SUBAPPLICATION Softkey_Aux_IXA_TO_Remote_WRITE_BG_Option_OPC (* VT-SoftKey lesen ODER AUX-Zuweisung (Joystick) lesen ODER lokaler Web-Override (z.B. vt-ui-mirror auf demselben Modul) + Remote-OPC-UA-Write an Zielmodul + VT-Hintergrundfarbe (SoftKey UND AUX) aus Remote-Subscribe - Option-Lib- Variante von Softkey_Aux_IXA_TO_Remote_WRITE_BG_OPC: Kommando-Seite komplett inaktiv (echtes INIT_REQ/INIT_CNF, kein VT-Object-Binding) wenn die Option nicht ausgewaehlt ist. Status-Seite (Remote-Subscribe) bleibt unveraendert immer aktiv - reiner Read ohne Seiteneffekt. *)
  (* Standard: 61499-2; Description: Copyright (c) 2026 Büngener Schuder GmbH This program and the accompanying materials are made available under the terms of the Eclipse Public License 2.0 which is available at https://www.eclipse.org/legal/epl-2.0/ SPDX-License-Identifier: EPL-2.0 *)
  (* Version 1.1, 2026-10-13, Franz Höpfinger, Büngener Schuder GmbH, Status jetzt auch Option-gated (AX_SUBSCRIBE_BG3_WEB_Option_OPC statt der ungated-Variante) - Franz: 'Command und STATUS muessen beide AUS/AN sein', 'reicht es alle Bausteine auszumachen die einen QI haben'. Command.PLUG1 -> Status.OPTION (sequenziell, Daisy-Chain analog OptionalGroup_001a/b) statt die Option-Socket zu splitten (strikt 1:1). Neuer eigener PLUG1-Ausgang reicht die Kette an weitere, dieselbe Option teilende Instanzen weiter (z.B. Bunker_Klappen_Auf -> Bunker_Klappen_Zu). *)
  (* Version 1.0, 2026-10-13, Franz Höpfinger, Büngener Schuder GmbH, initial implementation (verworfen, siehe v1.1) - duennwandiger Wrapper analog Softkey_Aux_IXA_TO_Remote_WRITE_BG_OPC, nutzt aber Softkey_Aux_IXA_TO_Remote_WRITE_Option (OPTION-Socket) statt der QI-Variante. Erster Aufrufer: Subscribe_STG3_Fanghaken (Franz: 'muss ein AOption Adapter sein'). *)
  PACKAGE MyLib::sys;
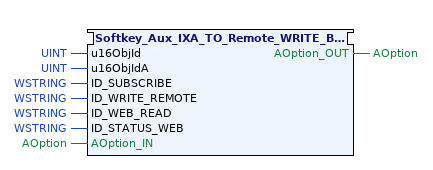
  VAR_INPUT
    u16ObjId : UINT; (* Object ID SoftKey/Hintergrund (VT) *)
    u16ObjIdA : UINT; (* Object ID AuxFunction2/Hintergrund (VT) *)
    ID_SUBSCRIBE : WSTRING; (* Remote-Subscribe-Adresse (Status/Farbe, ACTION=SUBSCRIBE) *)
    ID_WRITE_REMOTE : WSTRING; (* Remote-Write-Adresse zum Zielmodul (Befehl, ACTION=WRITE, CLIENT) *)
    ID_WEB_READ : WSTRING; (* Lokale Subscribe-Adresse fuer einen Web-Client (z.B. vt-ui-mirror) auf demselben Modul, ODER-verknuepft mit SoftKey und AUX *)
    ID_STATUS_WEB : WSTRING; (* Lokale Publish-Adresse (auf diesem Modul) fuer den vom Zielmodul zurueckgemeldeten Zustand - damit ein Web-Client (z.B. vt-ui-mirror) dieselbe Hintergrundfarbe wie das echte VT zeigen kann *)
  END_VAR
  SOCKETS
    AOption_IN : Option::AOption; (* Treibt INIT/QI von Command UND Status sequenziell - anschliessen an z.B. AOption_AUI_DEMUX_N.OUTx oder das PLUG1 einer vorgeschalteten Instanz *)
  END_SOCKETS
  PLUGS
    AOption_OUT : Option::AOption; (* Reicht die Aktivierung an eine nachgeschaltete Instanz weiter (Daisy-Chain, z.B. eine 2. SoftKey_Aux_IXA_TO_Remote_WRITE_BG_Option_OPC-Instanz, die dieselbe Option teilt) - unbenutzt lassen, wenn nichts weiter folgt *)
  END_PLUGS
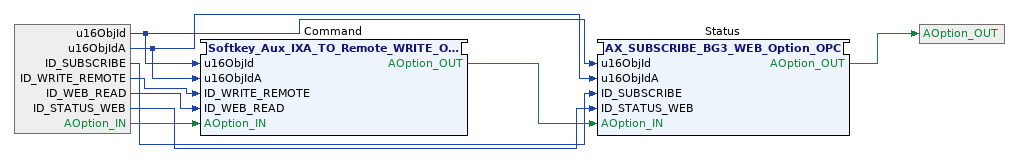
  SUBAPPS
    Command : MyLib::sys::Softkey_Aux_IXA_TO_Remote_WRITE_Option;
    Status : MyLib::sys::AX_SUBSCRIBE_BG3_WEB_Option_OPC;
  END_SUBAPPS
  DATA_CONNECTIONS
    u16ObjId TO Command.u16ObjId;
    u16ObjIdA TO Command.u16ObjIdA;
    ID_WRITE_REMOTE TO Command.ID_WRITE_REMOTE;
    ID_WEB_READ TO Command.ID_WEB_READ;
    u16ObjId TO Status.u16ObjId;
    u16ObjIdA TO Status.u16ObjIdA;
    ID_SUBSCRIBE TO Status.ID_SUBSCRIBE;
    ID_STATUS_WEB TO Status.ID_STATUS_WEB;
  END_CONNECTIONS
  ADAPTER_CONNECTIONS
    Command.AOption_OUT TO Status.AOption_IN;
    Status.AOption_OUT TO AOption_OUT;
    AOption_IN TO Command.AOption_IN;
  END_CONNECTIONS
END_SUBAPPLICATION
